(* IEC 61131-3 sources: GenAI/codesys_service/bank/st, 20 files *)

(* ---- E01_Filling.st ---- *)
FUNCTION_BLOCK E01_Filling
VAR_INPUT
    bottleSensor : BOOL;
    cleaningConfirmButton : BOOL;
    fillingConfirmButton : BOOL;
    cappingConfirmButton : BOOL;
    packingConfirmButton : BOOL;
    finishedButton : BOOL;
END_VAR
VAR_OUTPUT
    Pump_Motor : BOOL;
    Filling_Valve : BOOL;
    Capping_Machine : BOOL;
    Packing_Machine : BOOL;
    Completion_Light : BOOL;
END_VAR
VAR
    step : INT;      (* 0=idle 1=cleaning 2=filling 3=capping 4=packing 5=done *)
    prevBottle : BOOL;
    prevCleaning : BOOL;
    prevFilling : BOOL;
    prevCapping : BOOL;
    prevPacking : BOOL;
    prevFinished : BOOL;
END_VAR

(* step transitions on rising edges *)
IF step = 0 AND bottleSensor AND NOT prevBottle THEN
    step := 1;
END_IF;
IF step = 1 AND cleaningConfirmButton AND NOT prevCleaning THEN
    step := 2;
END_IF;
IF step = 2 AND fillingConfirmButton AND NOT prevFilling THEN
    step := 3;
END_IF;
IF step = 3 AND cappingConfirmButton AND NOT prevCapping THEN
    step := 4;
END_IF;
IF step = 4 AND packingConfirmButton AND NOT prevPacking THEN
    step := 5;
END_IF;
IF step = 5 AND finishedButton AND NOT prevFinished THEN
    step := 0;
END_IF;

(* outputs by step *)
Pump_Motor := (step = 1);
Filling_Valve := (step = 2);
Capping_Machine := (step = 3);
Packing_Machine := (step = 4);
Completion_Light := (step = 5);

prevBottle := bottleSensor;
prevCleaning := cleaningConfirmButton;
prevFilling := fillingConfirmButton;
prevCapping := cappingConfirmButton;
prevPacking := packingConfirmButton;
prevFinished := finishedButton;

(* ---- E02_DualEdge.st ---- *)
FUNCTION_BLOCK E02_DualEdge
VAR_INPUT
    value : DWORD;
END_VAR
VAR_OUTPUT
    hasChanged : BOOL;
    hasRisingEdges : BOOL;
    risingBits : DWORD;
    noOfRisingBits : USINT;
    hasFallingEdges : BOOL;
    fallingBits : DWORD;
    noOfFallingBits : USINT;
END_VAR
VAR
    prevValue : DWORD;
    i : INT;
    tr : DWORD;
    tf : DWORD;
    cntR : USINT;
    cntF : USINT;
END_VAR

risingBits := value AND (NOT prevValue);
fallingBits := (NOT value) AND prevValue;
hasChanged := (value <> prevValue);
hasRisingEdges := (risingBits <> 0);
hasFallingEdges := (fallingBits <> 0);

(* popcount without SHL: shift right by division *)
cntR := 0;
tr := risingBits;
FOR i := 0 TO 31 DO
    IF (tr MOD 2) = 1 THEN
        cntR := cntR + 1;
    END_IF;
    tr := tr / 2;
END_FOR;

cntF := 0;
tf := fallingBits;
FOR i := 0 TO 31 DO
    IF (tf MOD 2) = 1 THEN
        cntF := cntF + 1;
    END_IF;
    tf := tf / 2;
END_FOR;

noOfRisingBits := cntR;
noOfFallingBits := cntF;
prevValue := value;

(* ---- E03_Hysteresis.st ---- *)
FUNCTION_BLOCK E03_Hysteresis
VAR_INPUT
    Value : REAL;
    hiLevel : REAL;
    loLevel : REAL;
    hystWindow : REAL;
END_VAR
VAR_OUTPUT
    hiAlarm : BOOL;
    loAlarm : BOOL;
    error : BOOL;
    status : WORD;
END_VAR

IF loLevel >= hiLevel THEN
    error := TRUE;
    status := 16#8001;
    hiAlarm := FALSE;
    loAlarm := FALSE;
ELSIF hystWindow >= (hiLevel - loLevel) THEN
    error := TRUE;
    status := 16#8002;
    hiAlarm := FALSE;
    loAlarm := FALSE;
ELSE
    error := FALSE;
    status := 16#0000;
    (* high alarm with hysteresis *)
    IF hiAlarm THEN
        IF Value < (hiLevel - hystWindow) THEN
            hiAlarm := FALSE;
        END_IF;
    ELSE
        IF Value > hiLevel THEN
            hiAlarm := TRUE;
        END_IF;
    END_IF;
    (* low alarm with hysteresis *)
    IF loAlarm THEN
        IF Value > (loLevel + hystWindow) THEN
            loAlarm := FALSE;
        END_IF;
    ELSE
        IF Value < loLevel THEN
            loAlarm := TRUE;
        END_IF;
    END_IF;
END_IF;

(* ---- E04_JamPump.st ---- *)
FUNCTION_BLOCK E04_JamPump
VAR_INPUT
    VISCOSITY_OK : BOOL;
    PASTE_E_STOP_NC : BOOL;
    DebounceTime : TIME;
    CycleTime : TIME;
END_VAR
VAR_OUTPUT
    VFD_RUN : BOOL;
    PUMP_MAINT_DUE : BOOL;
    PUMP_RUNTIME_ACC : LTIME;
END_VAR
VAR
    viscTimer : TON;
    viscValid : BOOL;
END_VAR

(* debounce: only counts while signal AND permissive are both TRUE,
   so an emergency stop clears incomplete timing immediately *)
viscTimer(IN := VISCOSITY_OK AND PASTE_E_STOP_NC, PT := DebounceTime);
viscValid := viscTimer.Q;

VFD_RUN := viscValid AND PASTE_E_STOP_NC;

IF VFD_RUN THEN
    PUMP_RUNTIME_ACC := PUMP_RUNTIME_ACC + TIME_TO_LTIME(CycleTime);
END_IF;

PUMP_MAINT_DUE := (PUMP_RUNTIME_ACC >= LTIME#500H);

(* ---- E05_WeldGap.st ---- *)
FUNCTION_BLOCK E05_WeldGap
VAR_INPUT
    Gap_Exceeded : BOOL;
    Weld_E_Stop_NC : BOOL;
    DebounceTime : TIME;
END_VAR
VAR_OUTPUT
    Operator_Alert : BOOL;
    Weld_Soft_Start_Active : BOOL;
END_VAR
VAR
    initTimer : TON;
    gapTimer : TON;
    initDone : BOOL;
END_VAR

(* 5s power-up inhibition; e-stop freezes it (IN=FALSE) *)
initTimer(IN := Weld_E_Stop_NC AND NOT initDone, PT := T#5S);
IF initTimer.Q THEN
    initDone := TRUE;
END_IF;

Weld_Soft_Start_Active := (NOT initDone) AND Weld_E_Stop_NC;

(* gap monitoring only after init, only while no e-stop;
   IN=FALSE on signal loss / e-stop clears the timing automatically *)
gapTimer(IN := Weld_E_Stop_NC AND initDone AND Gap_Exceeded, PT := DebounceTime);
Operator_Alert := gapTimer.Q AND Weld_E_Stop_NC AND initDone;

(* ---- E06_Blower.st ---- *)
FUNCTION_BLOCK E06_Blower
VAR_INPUT
    DO_LOW : BOOL;
    AERATION_E_STOP_NC : BOOL;
END_VAR
VAR_OUTPUT
    BLOWER_RUN : BOOL;
    AERATION_BLOWER_CYCLE_COUNT : UINT;
END_VAR
VAR
    delayTimer : TON;
    prevRun : BOOL;
END_VAR

(* 5s start delay: IN goes FALSE on demand loss or e-stop, resetting timing *)
delayTimer(IN := DO_LOW AND AERATION_E_STOP_NC, PT := T#5S);
BLOWER_RUN := delayTimer.Q;

IF BLOWER_RUN AND NOT prevRun THEN
    AERATION_BLOWER_CYCLE_COUNT := AERATION_BLOWER_CYCLE_COUNT + 1;
END_IF;
prevRun := BLOWER_RUN;

(* ---- H01_Proportion.st ---- *)
FUNCTION_BLOCK H01_Proportion
VAR_INPUT
    estop : BOOL;
    opeMode : BOOL;
    valveAStart : BOOL;
    valveBStart : BOOL;
    valveCStart : BOOL;
    valveDStart : BOOL;
    mixMotorStart : BOOL;
    autoStart : BOOL;
    processMode : BOOL;
    levelSensor : INT;
    mixMotorComplete : BOOL;
END_VAR
VAR_OUTPUT
    valveARun : BOOL;
    valveBRun : BOOL;
    valveCRun : BOOL;
    valveDRun : BOOL;
    mixMotorRun : BOOL;
END_VAR
VAR
    step : INT;  (* 0=idle 1=fillA 2=fillB 3=fillC 4=mixing 5=done *)
    prevAuto : BOOL;
    prevVA : BOOL;
    prevVB : BOOL;
    prevVC : BOOL;
    prevVD : BOOL;
    prevMix : BOOL;
END_VAR

IF NOT estop THEN
    (* emergency stop: everything off, sequence aborted *)
    valveARun := FALSE;
    valveBRun := FALSE;
    valveCRun := FALSE;
    valveDRun := FALSE;
    mixMotorRun := FALSE;
    step := 0;
ELSIF NOT opeMode THEN
    (* manual mode: each button toggles its device on a rising edge *)
    IF valveAStart AND NOT prevVA THEN
        valveARun := NOT valveARun;
    END_IF;
    IF valveBStart AND NOT prevVB THEN
        valveBRun := NOT valveBRun;
    END_IF;
    IF valveCStart AND NOT prevVC THEN
        valveCRun := NOT valveCRun;
    END_IF;
    IF valveDStart AND NOT prevVD THEN
        valveDRun := NOT valveDRun;
    END_IF;
    IF mixMotorStart AND NOT prevMix THEN
        mixMotorRun := NOT mixMotorRun;
    END_IF;
    step := 0;
ELSE
    (* automatic mode state machine *)
    valveCRun := FALSE;
    mixMotorRun := FALSE;
    IF step = 0 THEN
        valveARun := FALSE;
        valveBRun := FALSE;
        valveDRun := FALSE;
        IF autoStart AND NOT prevAuto THEN
            valveARun := TRUE;
            step := 1;
        END_IF;
    ELSIF step = 1 THEN
        valveARun := TRUE;
        IF levelSensor >= 50 THEN
            valveARun := FALSE;
            valveBRun := TRUE;
            step := 2;
        END_IF;
    ELSIF step = 2 THEN
        valveBRun := TRUE;
        IF levelSensor >= 80 THEN
            valveBRun := FALSE;
            IF processMode THEN
                valveCRun := TRUE;
                step := 3;
            ELSE
                mixMotorRun := TRUE;
                step := 4;
            END_IF;
        END_IF;
    ELSIF step = 3 THEN
        valveCRun := TRUE;
        IF levelSensor >= 100 THEN
            valveCRun := FALSE;
            mixMotorRun := TRUE;
            step := 4;
        END_IF;
    ELSIF step = 4 THEN
        mixMotorRun := TRUE;
        IF mixMotorComplete THEN
            mixMotorRun := FALSE;
            valveDRun := TRUE;
            step := 5;
        END_IF;
    ELSE
        (* step 5: process finished, valve D stays open *)
        valveDRun := TRUE;
    END_IF;
END_IF;

prevAuto := autoStart;
prevVA := valveAStart;
prevVB := valveBStart;
prevVC := valveCStart;
prevVD := valveDStart;
prevMix := mixMotorStart;

(* ---- H02_FlexProcess.st ---- *)
FUNCTION_BLOCK H02_FlexProcess
VAR_INPUT
    processLength : USINT;
    sensor1 : BOOL;
    sensor2 : BOOL;
    sensor3 : BOOL;
    sensor4 : BOOL;
    sensor5 : BOOL;
    station1Start : BOOL;
    station2Complete : BOOL;
    station3Complete : BOOL;
    station4Complete : BOOL;
    processSequence : ARRAY[1..8] OF USINT;
END_VAR
VAR_OUTPUT
    conveyorLeft : BOOL;
    conveyorRight : BOOL;
END_VAR
VAR
    idx : INT := 1;      (* next sequence entry to execute *)
    cur : INT := 1;      (* current station position *)
    tgt : INT;           (* target station *)
    moving : BOOL;
    prevStart : BOOL;
    done : BOOL;
END_VAR

conveyorLeft := FALSE;
conveyorRight := FALSE;

IF (idx > processLength) OR (processLength < 1) OR (processLength > 8) THEN
    (* sequence exhausted: stay idle *)
    moving := FALSE;
    done := (idx > processLength) AND (processLength >= 1);
ELSE
    tgt := processSequence[idx];

    IF NOT moving THEN
        done := FALSE;
        IF cur = 1 THEN
            (* waiting at loading station for start *)
            IF sensor1 AND station1Start AND NOT prevStart THEN
                moving := TRUE;
            END_IF;
        ELSE
            (* waiting for completion signal of the current processing station *)
            IF (cur = 2 AND station2Complete)
                OR (cur = 3 AND station3Complete)
                OR (cur = 4 AND station4Complete) THEN
                moving := TRUE;
            END_IF;
        END_IF;
    END_IF;

    IF moving THEN
        IF tgt > cur THEN
            conveyorRight := TRUE;
        ELSIF tgt < cur THEN
            conveyorLeft := TRUE;
        END_IF;
        (* stop on arrival at the target station *)
        IF (tgt = 2 AND sensor2)
            OR (tgt = 3 AND sensor3)
            OR (tgt = 4 AND sensor4)
            OR (tgt = 5 AND sensor5) THEN
            moving := FALSE;
            conveyorLeft := FALSE;
            conveyorRight := FALSE;
            cur := tgt;
            idx := idx + 1;
        END_IF;
    END_IF;
END_IF;

prevStart := station1Start;

(* ---- H03_RecipeMgr.st ---- *)
TYPE ST_Recipe :
STRUCT
    recipeID : INT;
    ingredientType : INT;
    ingredientRatio : REAL;
    productionTemperature : REAL;
END_STRUCT
END_TYPE

FUNCTION_BLOCK H03_RecipeMgr
VAR_INPUT
    addRecipe : BOOL;
    deleteRecipe : BOOL;
    modifyRecipe : BOOL;
    queryRecipe : BOOL;
    recipeIn : ST_Recipe;
END_VAR
VAR_OUTPUT
    recipeAdded : BOOL;
    recipeDeleted : BOOL;
    recipeModified : BOOL;
    recipeQueryResult : ST_Recipe;
    error : BOOL;
    status : WORD;
END_VAR
VAR_IN_OUT
    recipe : ARRAY[1..10] OF ST_Recipe;
END_VAR
VAR
    i : INT;
    found : INT;
    freeSlot : INT;
    prevAdd : BOOL;
    prevDelete : BOOL;
    prevModify : BOOL;
    prevQuery : BOOL;
END_VAR

recipeAdded := FALSE;
recipeDeleted := FALSE;
recipeModified := FALSE;
error := FALSE;
status := 16#0000;
recipeQueryResult.recipeID := 0;
recipeQueryResult.ingredientType := 0;
recipeQueryResult.ingredientRatio := 0.0;
recipeQueryResult.productionTemperature := 0.0;

IF queryRecipe AND NOT prevQuery THEN
    found := 0;
    FOR i := 1 TO 10 DO
        IF recipe[i].recipeID = recipeIn.recipeID THEN
            found := i;
        END_IF;
    END_FOR;
    IF found = 0 THEN
        error := TRUE;
        status := 16#8001;
    ELSE
        recipeQueryResult := recipe[found];
    END_IF;

ELSIF addRecipe AND NOT prevAdd THEN
    found := 0;
    freeSlot := 0;
    FOR i := 1 TO 10 DO
        IF recipe[i].recipeID = recipeIn.recipeID THEN
            found := i;
        END_IF;
        IF (freeSlot = 0) AND (recipe[i].recipeID = 0) THEN
            freeSlot := i;
        END_IF;
    END_FOR;
    IF found <> 0 THEN
        error := TRUE;
        status := 16#8002;
    ELSIF freeSlot = 0 THEN
        error := TRUE;
        status := 16#8003;
    ELSE
        recipe[freeSlot] := recipeIn;
        recipeAdded := TRUE;
    END_IF;

ELSIF deleteRecipe AND NOT prevDelete THEN
    found := 0;
    FOR i := 1 TO 10 DO
        IF recipe[i].recipeID = recipeIn.recipeID THEN
            found := i;
        END_IF;
    END_FOR;
    IF found = 0 THEN
        error := TRUE;
        status := 16#8004;
    ELSE
        recipe[found].recipeID := 0;
        recipeDeleted := TRUE;
    END_IF;

ELSIF modifyRecipe AND NOT prevModify THEN
    found := 0;
    FOR i := 1 TO 10 DO
        IF recipe[i].recipeID = recipeIn.recipeID THEN
            found := i;
        END_IF;
    END_FOR;
    IF found = 0 THEN
        error := TRUE;
        status := 16#8005;
    ELSE
        recipe[found] := recipeIn;
        recipeModified := TRUE;
    END_IF;
END_IF;

prevAdd := addRecipe;
prevDelete := deleteRecipe;
prevModify := modifyRecipe;
prevQuery := queryRecipe;

(* ---- H04_FIFO.st ---- *)
(* 题面要求 item/buffer 为 VARIANT；纯 ST 无法对 VARIANT 做下标访问，
   此参考实现固定为 DINT / ARRAY[0..7] OF DINT 以验证逻辑，编译侧
   VARIANT 绑定能力另行验证。 *)
FUNCTION_BLOCK H04_FIFO
VAR_INPUT
    enqueue : BOOL;
    dequeue : BOOL;
    reset : BOOL;
END_VAR
VAR_OUTPUT
    elementCount : DINT;
    status : WORD;
END_VAR
VAR_IN_OUT
    item : DINT;
    buffer : ARRAY[0..7] OF DINT;
END_VAR
VAR
    head : DINT := 0;
    tail : DINT := 0;
    nq : DINT := 0;
    prevEnq : BOOL;
    prevDeq : BOOL;
    enqEdge : BOOL;
    deqEdge : BOOL;
END_VAR

IF reset THEN
    head := 0;
    tail := 0;
    nq := 0;
    elementCount := 0;
    status := 16#0000;
ELSE
    status := 16#0000;
    enqEdge := enqueue AND NOT prevEnq;
    deqEdge := dequeue AND NOT prevDeq;

    IF deqEdge THEN
        IF nq = 0 THEN
            status := 16#8001;   (* dequeue on empty queue *)
        ELSE
            item := buffer[head];
            head := head + 1;
            IF head > 7 THEN
                head := 0;
            END_IF;
            nq := nq - 1;
        END_IF;
    ELSIF enqEdge THEN
        IF nq >= 8 THEN
            status := 16#8002;   (* enqueue on full queue *)
        ELSE
            buffer[tail] := item;
            tail := tail + 1;
            IF tail > 7 THEN
                tail := 0;
            END_IF;
            nq := nq + 1;
        END_IF;
    END_IF;
    elementCount := nq;
END_IF;

prevEnq := enqueue;
prevDeq := dequeue;

(* ---- H05_MechArm.st ---- *)
FUNCTION_BLOCK H05_MechArm
VAR_INPUT
    ManualMode : BOOL;
    SingleStepMode : BOOL;
    SingleCycleMode : BOOL;
    ContinuousMode : BOOL;
    EmergencyStop : BOOL;
    Start : BOOL;
    DownButton : BOOL;
    UpButton : BOOL;
    LeftButton : BOOL;
    RightButton : BOOL;
    GripButton : BOOL;
    ReleaseButton : BOOL;
    DownLimitSwitch : BOOL;
    UpLimitSwitch : BOOL;
    LeftLimitSwitch : BOOL;
    RightLimitSwitch : BOOL;
    GripLimitSwitch : BOOL;
    ReleaseLimitSwitch : BOOL;
END_VAR
VAR_OUTPUT
    MoveDown : BOOL;
    MoveUp : BOOL;
    MoveLeft : BOOL;
    MoveRight : BOOL;
    ActivateGrip : BOOL;
    ActivateRelease : BOOL;
END_VAR
VAR
    step : INT := 0;   (* 0 idle, then 1..8 = the 8-action cycle *)
    prevStart : BOOL;
    running : BOOL;
END_VAR

MoveDown := FALSE;
MoveUp := FALSE;
MoveLeft := FALSE;
MoveRight := FALSE;
ActivateGrip := FALSE;
ActivateRelease := FALSE;

IF NOT EmergencyStop THEN
    (* emergency stop: all actions off, sequence aborted *)
    step := 0;
    running := FALSE;
ELSIF ManualMode THEN
    (* manual: buttons drive actions, limited by position switches *)
    MoveDown := DownButton AND NOT DownLimitSwitch;
    MoveUp := UpButton AND NOT UpLimitSwitch;
    MoveLeft := LeftButton AND NOT LeftLimitSwitch;
    MoveRight := RightButton AND NOT RightLimitSwitch;
    ActivateGrip := GripButton AND NOT GripLimitSwitch;
    ActivateRelease := ReleaseButton AND NOT ReleaseLimitSwitch;
    step := 0;
    running := FALSE;
ELSIF SingleStepMode THEN
    (* single step: each start press advances one action *)
    IF Start AND NOT prevStart AND NOT running THEN
        IF step = 0 THEN
            step := 1;
        END_IF;
    END_IF;
    IF step > 0 THEN
        running := TRUE;
    END_IF;
ELSE
    (* single cycle / continuous: run through the cycle automatically *)
    IF (Start AND NOT prevStart) AND (step = 0) THEN
        step := 1;
    END_IF;
    IF step > 0 THEN
        running := TRUE;
    END_IF;
END_IF;

IF running AND EmergencyStop THEN
    (* action execution by step; each step stops on its completion feedback *)
    IF step = 1 THEN
        MoveDown := NOT DownLimitSwitch;
        IF DownLimitSwitch THEN step := 2; END_IF;
    ELSIF step = 2 THEN
        ActivateGrip := NOT GripLimitSwitch;
        IF GripLimitSwitch THEN step := 3; END_IF;
    ELSIF step = 3 THEN
        MoveUp := NOT UpLimitSwitch;
        IF UpLimitSwitch THEN step := 4; END_IF;
    ELSIF step = 4 THEN
        MoveRight := NOT RightLimitSwitch;
        IF RightLimitSwitch THEN step := 5; END_IF;
    ELSIF step = 5 THEN
        MoveDown := NOT DownLimitSwitch;
        IF DownLimitSwitch THEN step := 6; END_IF;
    ELSIF step = 6 THEN
        ActivateRelease := NOT ReleaseLimitSwitch;
        IF ReleaseLimitSwitch THEN step := 7; END_IF;
    ELSIF step = 7 THEN
        MoveUp := NOT UpLimitSwitch;
        IF UpLimitSwitch THEN step := 8; END_IF;
    ELSIF step = 8 THEN
        MoveLeft := NOT LeftLimitSwitch;
        IF LeftLimitSwitch THEN
            (* cycle complete: single cycle stops, continuous restarts *)
            IF ContinuousMode THEN
                step := 1;
            ELSE
                step := 0;
                running := FALSE;
            END_IF;
        END_IF;
    ELSE
        running := FALSE;
    END_IF;

    (* single step pauses between actions after completing one *)
    IF SingleStepMode AND (step > 1) THEN
        (* stop execution after the current action finishes:
           handled implicitly on the next invocation *)
        running := FALSE;
        step := step;  (* hold position, wait for next start *)
    END_IF;
END_IF;

prevStart := Start;

(* ---- H06_Production.st ---- *)
FUNCTION_BLOCK H06_Production
VAR_INPUT
    Mode : BOOL;
    ForwardButton : BOOL;
    ReverseButton : BOOL;
    SensorFeed : BOOL;
    SensorWash : BOOL;
    SensorWeight : BOOL;
    SensorFiring : BOOL;
    SensorOutput : BOOL;
    washComplete : BOOL;
    weightComplete : BOOL;
    weight : REAL;
    firingComplete : BOOL;
END_VAR
VAR_OUTPUT
    MotorForward : BOOL;
    MotorReverse : BOOL;
    kick : BOOL;
    CompletionLight : BOOL;
    firingTemp : REAL;
END_VAR
VAR
    step : INT;  (* 0=feed 1=feed->wash 2=wash wait 3=wash->weight 4=weigh
                    5=weight->(kick|fire) 6=fire wait 7=fire->out 8=done *)
    qualified : BOOL;
    prevWashC : BOOL;
    prevWeightC : BOOL;
    prevFireC : BOOL;
END_VAR

IF NOT Mode THEN
    MotorForward := ForwardButton AND NOT ReverseButton;
    MotorReverse := ReverseButton AND NOT ForwardButton;
    kick := FALSE;
    CompletionLight := FALSE;
    step := 0;
ELSE
    MotorReverse := FALSE;
    IF step = 0 THEN
        MotorForward := FALSE;
        kick := FALSE;
        IF SensorFeed THEN
            step := 1;
        END_IF;
    ELSIF step = 1 THEN
        MotorForward := TRUE;
        IF SensorWash THEN
            MotorForward := FALSE;
            step := 2;
        END_IF;
    ELSIF step = 2 THEN
        MotorForward := FALSE;
        IF washComplete AND NOT prevWashC THEN
            step := 3;
        END_IF;
    ELSIF step = 3 THEN
        MotorForward := TRUE;
        IF SensorWeight THEN
            MotorForward := FALSE;
            step := 4;
        END_IF;
    ELSIF step = 4 THEN
        MotorForward := FALSE;
        IF weightComplete AND NOT prevWeightC THEN
            qualified := (weight >= 100.0) AND (weight <= 200.0);
            IF qualified THEN
                (* 100..200 kg -> 500..550 degrees, linear *)
                firingTemp := 500.0 + (weight - 100.0) * 0.5;
                step := 5;
            ELSE
                kick := TRUE;
                step := 8;
            END_IF;
        END_IF;
    ELSIF step = 5 THEN
        MotorForward := TRUE;
        IF SensorFiring THEN
            MotorForward := FALSE;
            step := 6;
        END_IF;
    ELSIF step = 6 THEN
        MotorForward := FALSE;
        IF firingComplete AND NOT prevFireC THEN
            step := 7;
        END_IF;
    ELSIF step = 7 THEN
        MotorForward := TRUE;
        IF SensorOutput THEN
            MotorForward := FALSE;
            step := 8;
        END_IF;
    ELSE
        (* step 8: finished / rejected *)
        MotorForward := FALSE;
        CompletionLight := SensorOutput;
        IF NOT SensorOutput THEN
            CompletionLight := FALSE;
            kick := FALSE;
            step := 0;
        END_IF;
    END_IF;
END_IF;

prevWashC := washComplete;
prevWeightC := weightComplete;
prevFireC := firingComplete;

(* ---- M01_PumpSwitch.st ---- *)
TYPE ST_Pump :
STRUCT
    priority : INT;
    selection : BOOL;
    RunComd : BOOL;
END_STRUCT
END_TYPE

FUNCTION_BLOCK M01_PumpSwitch
VAR_INPUT
    mode : BOOL;
    start : BOOL;
    stop : BOOL;
END_VAR
VAR_IN_OUT
    pumpGroup : ARRAY[1..5] OF ST_Pump;
END_VAR
VAR_OUTPUT
    runningCount : INT;
END_VAR
VAR
    i : INT;
    j : INT;
    rank : INT;
END_VAR

IF stop THEN
    FOR i := 1 TO 5 DO
        pumpGroup[i].RunComd := FALSE;
    END_FOR;
ELSIF mode THEN
    (* automatic: rank by priority, ties broken by index; top 3 run *)
    FOR i := 1 TO 5 DO
        rank := 1;
        FOR j := 1 TO 5 DO
            IF j <> i THEN
                IF (pumpGroup[j].priority > pumpGroup[i].priority)
                    OR ((pumpGroup[j].priority = pumpGroup[i].priority) AND (j < i)) THEN
                    rank := rank + 1;
                END_IF;
            END_IF;
        END_FOR;
        pumpGroup[i].RunComd := start AND (rank <= 3);
    END_FOR;
ELSE
    (* manual: selected pumps start with the start button *)
    FOR i := 1 TO 5 DO
        pumpGroup[i].RunComd := start AND pumpGroup[i].selection;
    END_FOR;
END_IF;

runningCount := 0;
FOR i := 1 TO 5 DO
    IF pumpGroup[i].RunComd THEN
        runningCount := runningCount + 1;
    END_IF;
END_FOR;

(* ---- M02_AnalogBatch.st ---- *)
TYPE ST_AnalogChannel :
STRUCT
    enable : BOOL;
    hiLIM : REAL;
    loLIM : REAL;
    bipolar : BOOL;
    measuringMode : INT;
    retVal : WORD;
    outputValue : REAL;
END_STRUCT
END_TYPE

FUNCTION_BLOCK M02_AnalogBatch
VAR_INPUT
    count : DINT;
END_VAR
VAR_IN_OUT
    analogValues : ARRAY[1..8] OF INT;
    channels : ARRAY[1..8] OF ST_AnalogChannel;
END_VAR
VAR
    k : DINT;
    raw : INT;
    ch : ST_AnalogChannel;
    res : REAL;
END_VAR

FOR k := 1 TO count DO
    IF channels[k].enable THEN
        raw := analogValues[k];
        IF channels[k].measuringMode = 0 THEN
            IF channels[k].hiLIM <= channels[k].loLIM THEN
                channels[k].retVal := 16#8002;
            ELSE
                IF channels[k].bipolar THEN
                    res := channels[k].loLIM
                           + (INT_TO_REAL(raw + 27648) / 55296.0)
                             * (channels[k].hiLIM - channels[k].loLIM);
                ELSE
                    res := channels[k].loLIM
                           + (INT_TO_REAL(raw) / 27648.0)
                             * (channels[k].hiLIM - channels[k].loLIM);
                END_IF;
                channels[k].outputValue := res;
                channels[k].retVal := 16#0000;
            END_IF;
        ELSIF channels[k].measuringMode = 1 THEN
            channels[k].outputValue := INT_TO_REAL(raw) / 10.0;
            channels[k].retVal := 16#0000;
        ELSIF channels[k].measuringMode = 2 THEN
            channels[k].outputValue := INT_TO_REAL(raw) / 100.0;
            channels[k].retVal := 16#0000;
        ELSE
            channels[k].retVal := 16#8001;
        END_IF;
    END_IF;
END_FOR;

(* ---- M03_MovingAvg.st ---- *)
FUNCTION_BLOCK M03_MovingAvg
VAR_INPUT
    cyclicExecution : BOOL;
    trigger : BOOL;
    value : LREAL;
    windowSize : INT;
    reset : BOOL;
END_VAR
VAR_OUTPUT
    average : LREAL;
    windowSizeReached : BOOL;
    error : BOOL;
    status : WORD;
END_VAR
VAR
    buf : ARRAY[1..100] OF LREAL;
    idx : INT := 1;
    filled : INT := 0;
    sum : LREAL := 0.0;
    prevTrigger : BOOL;
    doUpdate : BOOL;
END_VAR

IF (windowSize < 1) OR (windowSize > 100) THEN
    error := TRUE;
    status := 16#8200;
    average := 0.0;
    windowSizeReached := FALSE;
ELSIF reset THEN
    filled := 0;
    idx := 1;
    sum := 0.0;
    average := 0.0;
    windowSizeReached := FALSE;
    error := FALSE;
    status := 16#0000;
ELSE
    error := FALSE;
    status := 16#0000;
    doUpdate := cyclicExecution OR (trigger AND NOT prevTrigger);
    IF doUpdate THEN
        IF filled < windowSize THEN
            (* filling phase: plain average of received values *)
            buf[idx] := value;
            sum := sum + value;
            filled := filled + 1;
            idx := idx + 1;
            IF idx > windowSize THEN
                idx := 1;
            END_IF;
            average := sum / INT_TO_LREAL(filled);
            windowSizeReached := (filled >= windowSize);
        ELSE
            (* steady state: replace oldest, recompute *)
            sum := sum - buf[idx] + value;
            buf[idx] := value;
            idx := idx + 1;
            IF idx > windowSize THEN
                idx := 1;
            END_IF;
            average := sum / INT_TO_LREAL(windowSize);
            windowSizeReached := TRUE;
        END_IF;
    END_IF;
END_IF;

prevTrigger := trigger;

(* ---- M04_TempCtrl.st ---- *)
FUNCTION_BLOCK M04_TempCtrl
VAR_INPUT
    TemperatureSensorInput : REAL;
    SetTemperature : REAL;
END_VAR
VAR_OUTPUT
    CurrentTemperature : REAL;
    SetTempDisplay : REAL;
    HeaterStatus : BOOL;
    OverheatProtection : BOOL;
    HeaterOutput : BOOL;
END_VAR
VAR
    heatTimer : TON;
    releaseTimer : TON;
    sensorFault : BOOL;
END_VAR

CurrentTemperature := TemperatureSensorInput;
SetTempDisplay := SetTemperature;

sensorFault := (TemperatureSensorInput < 0.0) OR (TemperatureSensorInput > 100.0);

IF sensorFault THEN
    HeaterOutput := FALSE;
    OverheatProtection := FALSE;
    heatTimer(IN := FALSE, PT := T#5S);
    releaseTimer(IN := FALSE, PT := T#3S);
ELSIF OverheatProtection THEN
    (* protection active: heater forced off, heat timing reset,
       lift after 3s pause *)
    HeaterOutput := FALSE;
    heatTimer(IN := FALSE, PT := T#5S);
    releaseTimer(IN := TRUE, PT := T#3S);
    IF releaseTimer.Q THEN
        OverheatProtection := FALSE;
    END_IF;
ELSE
    HeaterOutput := (TemperatureSensorInput < SetTemperature);
    heatTimer(IN := HeaterOutput, PT := T#5S);
    releaseTimer(IN := FALSE, PT := T#3S);
    IF heatTimer.Q THEN
        OverheatProtection := TRUE;
        HeaterOutput := FALSE;
    END_IF;
END_IF;

HeaterStatus := HeaterOutput;

(* ---- M05_ProdLine.st ---- *)
FUNCTION_BLOCK M05_ProdLine
VAR_INPUT
    Mode : BOOL;
    ForwardButton : BOOL;
    ReverseButton : BOOL;
    SensorA : BOOL;
    SensorB : BOOL;
    SensorC : BOOL;
    ButtonA : BOOL;
    ButtonB : BOOL;
    ButtonC : BOOL;
END_VAR
VAR_OUTPUT
    MotorForward : BOOL;
    MotorReverse : BOOL;
    CompletionLight : BOOL;
END_VAR
VAR
    step : INT;   (* 0=at A waiting 1=A->B 2=at B waiting 3=B->C 4=at C done *)
    prevA : BOOL;
    prevB : BOOL;
    prevC : BOOL;
END_VAR

IF NOT Mode THEN
    (* manual mode with forward/reverse interlock *)
    MotorForward := ForwardButton AND NOT ReverseButton;
    MotorReverse := ReverseButton AND NOT ForwardButton;
    CompletionLight := FALSE;
ELSE
    MotorReverse := FALSE;
    IF step = 0 THEN
        MotorForward := FALSE;
        IF SensorA AND ButtonA AND NOT prevA THEN
            step := 1;
        END_IF;
    ELSIF step = 1 THEN
        MotorForward := TRUE;
        IF SensorB THEN
            MotorForward := FALSE;
            step := 2;
        END_IF;
    ELSIF step = 2 THEN
        MotorForward := FALSE;
        IF ButtonB AND NOT prevB THEN
            step := 3;
        END_IF;
    ELSIF step = 3 THEN
        MotorForward := TRUE;
        IF SensorC THEN
            MotorForward := FALSE;
            step := 4;
        END_IF;
    ELSE
        (* step 4: at C *)
        MotorForward := FALSE;
        IF ButtonC AND NOT prevC THEN
            CompletionLight := TRUE;
        END_IF;
        IF NOT SensorC THEN
            CompletionLight := FALSE;
            step := 0;
        END_IF;
    END_IF;
END_IF;

prevA := ButtonA;
prevB := ButtonB;
prevC := ButtonC;

(* ---- M06_SlabThick.st ---- *)
FUNCTION_BLOCK M06_SlabThick
VAR_INPUT
    THICKNESS_FAULT : BOOL;
    THICKNESS_SIGNAL_VALID : BOOL;
    CUTTING_RUN : BOOL;
    FaultTimestamp : DINT;
    CycleTime : TIME;
END_VAR
VAR_OUTPUT
    THICKNESS_ALARM : BOOL;
    Slab_Fault_Counter : UINT;
    Slab_Runtime_Accumulator : LTIME;
    Slab_Fault_History : ARRAY[0..4] OF DINT;
END_VAR
VAR
    holdTimer : TOF;
    prevFault : BOOL;
END_VAR

IF THICKNESS_SIGNAL_VALID THEN
    (* alarm with minimum 500ms hold (TOF) while fault persists *)
    holdTimer(IN := THICKNESS_FAULT, PT := T#500MS);
    THICKNESS_ALARM := THICKNESS_FAULT OR holdTimer.Q;

    (* fault bookkeeping on rising edge of a valid fault *)
    IF THICKNESS_FAULT AND NOT prevFault THEN
        Slab_Fault_Counter := Slab_Fault_Counter + 1;
        Slab_Fault_History[4] := Slab_Fault_History[3];
        Slab_Fault_History[3] := Slab_Fault_History[2];
        Slab_Fault_History[2] := Slab_Fault_History[1];
        Slab_Fault_History[1] := Slab_Fault_History[0];
        Slab_Fault_History[0] := FaultTimestamp;
    END_IF;

    (* normal-cutting runtime accumulation *)
    IF CUTTING_RUN AND NOT THICKNESS_FAULT THEN
        Slab_Runtime_Accumulator := Slab_Runtime_Accumulator + TIME_TO_LTIME(CycleTime);
    END_IF;
ELSE
    (* signal invalid: alarm off, holding state cleared *)
    THICKNESS_ALARM := FALSE;
    holdTimer(IN := FALSE, PT := T#500MS);
END_IF;

prevFault := THICKNESS_FAULT;

(* ---- M07_HVAC.st ---- *)
FUNCTION_BLOCK M07_HVAC
VAR_INPUT
    OCCUPANCY_DETECTED : BOOL;
    ENERGY_SAVING_MODE : BOOL;
    HVAC_MODE_SELECTOR : INT;
END_VAR
VAR_OUTPUT
    SUPPLY_FAN_RUN : BOOL;
    TEMP_SETPOINT_ADJUST : INT;
END_VAR
VAR
    fanDelay : TON;
END_VAR

(* 30s start delay: any condition loss resets timing *)
fanDelay(IN := OCCUPANCY_DETECTED AND (HVAC_MODE_SELECTOR <> 3), PT := T#30S);
SUPPLY_FAN_RUN := fanDelay.Q;

IF HVAC_MODE_SELECTOR = 0 THEN
    (* Auto *)
    IF OCCUPANCY_DETECTED THEN
        TEMP_SETPOINT_ADJUST := 0;
    ELSIF ENERGY_SAVING_MODE THEN
        TEMP_SETPOINT_ADJUST := 3;
    ELSE
        TEMP_SETPOINT_ADJUST := 2;
    END_IF;
ELSIF HVAC_MODE_SELECTOR = 1 THEN
    (* Comfort *)
    IF OCCUPANCY_DETECTED THEN
        TEMP_SETPOINT_ADJUST := 0;
    ELSE
        TEMP_SETPOINT_ADJUST := 1;
    END_IF;
ELSIF HVAC_MODE_SELECTOR = 2 THEN
    (* Economy *)
    IF OCCUPANCY_DETECTED THEN
        TEMP_SETPOINT_ADJUST := 0;
    ELSE
        TEMP_SETPOINT_ADJUST := 4;
    END_IF;
ELSE
    (* Night *)
    TEMP_SETPOINT_ADJUST := 4;
END_IF;

(* ---- M08_IPv4.st ---- *)
FUNCTION_BLOCK M08_IPv4
VAR_INPUT
    ipText : STRING(254);
END_VAR
VAR_OUTPUT
    ipValue : UDINT;
END_VAR
VAR
    i : INT;
    ch : BYTE;
    seg : DINT;
    segCount : INT;
    started : BOOL;
    ok : BOOL;
    acc : DINT;
    slen : INT;
END_VAR

(* Standard Library: LEN gives the number of characters; the STRING itself
   is indexed directly (1-based) to avoid repeated MID copies. *)
ipValue := 0;
ok := TRUE;
seg := 0;
segCount := 0;
started := FALSE;
acc := 0;
slen := LEN(ipText);

FOR i := 1 TO slen DO
    ch := ipText[i];
    IF ch = 46 THEN
        (* '.' separator *)
        IF (NOT started) OR (seg > 255) OR (segCount = 4) THEN
            ok := FALSE;
        ELSE
            acc := acc * 256 + seg;
            segCount := segCount + 1;
            seg := 0;
            started := FALSE;
        END_IF;
    ELSIF (ch >= 48) AND (ch <= 57) THEN
        (* decimal digit *)
        seg := seg * 10 + (ch - 48);
        started := TRUE;
    ELSE
        ok := FALSE;
    END_IF;
END_FOR;

(* final segment must be present and in range; exactly 4 segments total *)
IF (NOT started) OR (seg > 255) OR (segCount <> 3) THEN
    ok := FALSE;
END_IF;

IF ok THEN
    acc := acc * 256 + seg;
    ipValue := DINT_TO_UDINT(acc);
ELSE
    ipValue := 0;
END_IF;
